{attribute 'qualified_only'}
{attribute 'strict'}
TYPE E_TankState :
(
	Idle	:= 0,
	Filling := 10,
	Full	:= 20,
	Draining := 30,
	Empty	:= 35,
	Manual	:= 40,
	Fault	:= 99
) INT;
END_TYPE

(* stored: Version 1.1.0.1
   DUT E_TankState: Id {c7aa19b8-0e8e-4367-99ba-0307db0aec77} *)
